// TIA Portal V19 export
DATA_BLOCK "Pumps Data"   // DB4
{ S7_Optimized_Access := 'FALSE'; DB_Accessible_From_OPC_UA := 'FALSE' }
// stored: DBAccessibleFromOPCUA false
   VAR RETAIN
      R1_CP01 : Struct
         MCMD : Bool;
         CMD : Bool;
         RESET : Bool;
         WT_SP : Time := T#5s;
         STATUS : Int;
      END_STRUCT;
      R1_AG01 : Struct
         MCMD : Bool;
         CMD : Bool;
         RESET : Bool;
         WT_SP : Time;
         STATUS : Int;
      END_STRUCT;
      CHS_CP01 : Struct
         MCMD : Bool;
         CMD : Bool;
         RESET : Bool;
         WT_SP : Time := T#5s;
         STATUS : Int;
         PUMP_SEL : Bool;
      END_STRUCT;
      CHS_CP02 : Struct
         MCMD : Bool;
         CMD : Bool;
         RESET : Bool;
         WT_SP : Time := T#5s;
         STATUS : Int;
         PUMP_SEL : Bool;
      END_STRUCT;
      CHS_CP03 : Struct
         MCMD : Bool;
         CMD : Bool;
         RESET : Bool;
         WT_SP : Time := T#5s;
         STATUS : Int;
         PUMP_SEL : Bool;
      END_STRUCT;
      R2_CP01 : Struct
         MCMD : Bool;
         CMD : Bool;
         RESET : Bool;
         WT_SP : Time := T#5s;
         STATUS : Int;
      END_STRUCT;
      R2_AG01 : Struct
         MCMD : Bool;
         CMD : Bool;
         RESET : Bool;
         WT_SP : Time;
         STATUS : Int;
      END_STRUCT;
      R3_CP01 : Struct
         MCMD : Bool;
         CMD : Bool;
         RESET : Bool;
         WT_SP : Time := T#5s;
         STATUS : Int;
      END_STRUCT;
      R3_AG01 : Struct
         MCMD : Bool;
         CMD : Bool;
         RESET : Bool;
         WT_SP : Time;
         STATUS : Int;
      END_STRUCT;
      R4_CP01 : Struct
         MCMD : Bool;
         CMD : Bool;
         RESET : Bool;
         WT_SP : Time := T#5s;
         STATUS : Int;
      END_STRUCT;
      R4_AG01 : Struct
         MCMD : Bool;
         CMD : Bool;
         RESET : Bool;
         WT_SP : Time;
         STATUS : Int;
      END_STRUCT;
      R5_CP01 : Struct
         MCMD : Bool;
         CMD : Bool;
         RESET : Bool;
         WT_SP : Time := T#5s;
         STATUS : Int;
      END_STRUCT;
      R5_AG01 : Struct
         MCMD : Bool;
         CMD : Bool;
         RESET : Bool;
         WT_SP : Time;
         STATUS : Int;
      END_STRUCT;
      R6_CP01 : Struct
         MCMD : Bool;
         CMD : Bool;
         RESET : Bool;
         WT_SP : Time := T#5s;
         STATUS : Int;
      END_STRUCT;
      R6_AG01 : Struct
         MCMD : Bool;
         CMD : Bool;
         RESET : Bool;
         WT_SP : Time;
         STATUS : Int;
      END_STRUCT;
      R7_CP01 : Struct
         MCMD : Bool;
         CMD : Bool;
         RESET : Bool;
         WT_SP : Time := T#5s;
         STATUS : Int;
      END_STRUCT;
      R7_AG01 : Struct
         MCMD : Bool;
         CMD : Bool;
         RESET : Bool;
         WT_SP : Time;
         STATUS : Int;
      END_STRUCT;
      R8_CP01 : Struct
         MCMD : Bool;
         CMD : Bool;
         RESET : Bool;
         WT_SP : Time := T#5s;
         STATUS : Int;
      END_STRUCT;
      R8_AG01 : Struct
         MCMD : Bool;
         CMD : Bool;
         RESET : Bool;
         WT_SP : Time;
         STATUS : Int;
      END_STRUCT;
      R9_CP01 : Struct
         MCMD : Bool;
         CMD : Bool;
         RESET : Bool;
         WT_SP : Time := T#5s;
         STATUS : Int;
      END_STRUCT;
      R9_AG01 : Struct
         MCMD : Bool;
         CMD : Bool;
         RESET : Bool;
         WT_SP : Time;
         STATUS : Int;
      END_STRUCT;
      R10_CP01 : Struct
         MCMD : Bool;
         CMD : Bool;
         RESET : Bool;
         WT_SP : Time := T#5s;
         STATUS : Int;
      END_STRUCT;
      R10_AG01 : Struct
         MCMD : Bool;
         CMD : Bool;
         RESET : Bool;
         WT_SP : Time;
         STATUS : Int;
      END_STRUCT;
      R11_CP01 : Struct
         MCMD : Bool;
         CMD : Bool;
         RESET : Bool;
         WT_SP : Time := T#5s;
         STATUS : Int;
      END_STRUCT;
      R11_AG01 : Struct
         MCMD : Bool;
         CMD : Bool;
         RESET : Bool;
         WT_SP : Time;
         STATUS : Int;
      END_STRUCT;
      R12_CP01 : Struct
         MCMD : Bool;
         CMD : Bool;
         RESET : Bool;
         WT_SP : Time := T#5s;
         STATUS : Int;
      END_STRUCT;
      R12_AG01 : Struct
         MCMD : Bool;
         CMD : Bool;
         RESET : Bool;
         WT_SP : Time;
         STATUS : Int;
      END_STRUCT;
      R13_CP01 : Struct
         MCMD : Bool;
         CMD : Bool;
         RESET : Bool;
         WT_SP : Time := T#5s;
         STATUS : Int;
      END_STRUCT;
      R13_AG01 : Struct
         MCMD : Bool;
         CMD : Bool;
         RESET : Bool;
         WT_SP : Time;
         STATUS : Int;
      END_STRUCT;
      R14_CP01 : Struct
         MCMD : Bool;
         CMD : Bool;
         RESET : Bool;
         WT_SP : Time := T#5s;
         STATUS : Int;
      END_STRUCT;
      R14_AG01 : Struct
         MCMD : Bool;
         CMD : Bool;
         RESET : Bool;
         WT_SP : Time;
         STATUS : Int;
      END_STRUCT;
      R15_CP01 : Struct
         MCMD : Bool;
         CMD : Bool;
         RESET : Bool;
         WT_SP : Time := T#5s;
         STATUS : Int;
      END_STRUCT;
      R15_AG01 : Struct
         MCMD : Bool;
         CMD : Bool;
         RESET : Bool;
         WT_SP : Time;
         STATUS : Int;
      END_STRUCT;
      R16_CP01 : Struct
         MCMD : Bool;
         CMD : Bool;
         RESET : Bool;
         WT_SP : Time := T#5s;
         STATUS : Int;
      END_STRUCT;
      R16_AG01 : Struct
         MCMD : Bool;
         CMD : Bool;
         RESET : Bool;
         WT_SP : Time;
         STATUS : Int;
      END_STRUCT;
      R17_CP01 : Struct
         MCMD : Bool;
         CMD : Bool;
         RESET : Bool;
         WT_SP : Time := T#5s;
         STATUS : Int;
      END_STRUCT;
      R17_AG01 : Struct
         MCMD : Bool;
         CMD : Bool;
         RESET : Bool;
         WT_SP : Time;
         STATUS : Int;
      END_STRUCT;
      R18_CP01 : Struct
         MCMD : Bool;
         CMD : Bool;
         RESET : Bool;
         WT_SP : Time := T#5s;
         STATUS : Int;
      END_STRUCT;
      R18_AG01 : Struct
         MCMD : Bool;
         CMD : Bool;
         RESET : Bool;
         WT_SP : Time;
         STATUS : Int;
      END_STRUCT;
      UCHS_CP01 : Struct
         MCMD : Bool;
         CMD : Bool;
         RESET : Bool;
         WT_SP : Time := T#5s;
         STATUS : Int;
         PUMP_SEL : Bool;
      END_STRUCT;
      UCHS_CP02 : Struct
         MCMD : Bool;
         CMD : Bool;
         RESET : Bool;
         WT_SP : Time := T#5s;
         STATUS : Int;
         PUMP_SEL : Bool;
      END_STRUCT;
      UCHS_PUPM_FAULT : Struct
         UCHS_CP01_FAIL_TO_RUN : Bool;
         UCHS_CP02_FAIL_TO_RUN : Bool;
         UCHS_CP03_FAIL_TO_RUN : Bool;
         UCHS_CP01_FAULTY : Bool;
         UCHS_CP02_FAULTY : Bool;
         UCHS_CP03_FAULTY : Bool;
      END_STRUCT;
      CS_CP01 : Struct
         MCMD : Bool;
         CMD : Bool;
         RESET : Bool;
         WT_SP : Time := T#5s;
         STATUS : Int;
         PUMP_SEL : Bool;
         "FAIL TO RUN" : Bool;
      END_STRUCT;
      CS_CP02 : Struct
         MCMD : Bool;
         CMD : Bool;
         RESET : Bool;
         WT_SP : Time := T#5s;
         STATUS : Int;
         PUMP_SEL : Bool;
         "FAIL TO RUN" : Bool;
      END_STRUCT;
      CS_CP03 : Struct
         MCMD : Bool;
         CMD : Bool;
         RESET : Bool;
         WT_SP : Time := T#5s;
         STATUS : Int;
         PUMP_SEL : Bool;
         "FAIL TO RUN" : Bool;
      END_STRUCT;
      CS_PUPM_FAULT : Struct
         CS_CP01_FAIL_TO_RUN : Bool;
         CS_CP02_FAIL_TO_RUN : Bool;
         CS_CP03_FAIL_TO_RUN : Bool;
         CS_CP01_FAULTY : Bool;
         CS_CP02_FAULTY : Bool;
         CS_CP03_FAULTY : Bool;
      END_STRUCT;
      HS_CP01 : Struct
         MCMD : Bool;
         CMD : Bool;
         RESET : Bool;
         WT_SP : Time := T#5s;
         STATUS : Int;
         PUMP_SEL : Bool;
      END_STRUCT;
      HS_CP02 : Struct
         MCMD : Bool;
         CMD : Bool;
         RESET : Bool;
         WT_SP : Time := T#5s;
         STATUS : Int;
         PUMP_SEL : Bool;
      END_STRUCT;
      HS_CP03 : Struct
         MCMD : Bool;
         CMD : Bool;
         RESET : Bool;
         WT_SP : Time := T#5s;
         STATUS : Int;
         PUMP_SEL : Bool;
      END_STRUCT;
      HS_PUPM_FAULT : Struct
         HS_CP01_FAIL_TO_RUN : Bool;
         HS_CP02_FAIL_TO_RUN : Bool;
         HS_CP03_FAIL_TO_RUN : Bool;
         HS_CP01_FAULTY : Bool;
         HS_CP02_FAULTY : Bool;
         HS_CP03_FAULTY : Bool;
      END_STRUCT;
      "A/SCRB_001_CP01" : Struct
         MCMD : Bool;
         CMD : Bool;
         RESET : Bool;
         WT_SP : Time := T#5s;
         STATUS : Int;
         PUMP_SEL : Bool;
      END_STRUCT;
      "A/SCRB_001_CP02" : Struct
         MCMD : Bool;
         CMD : Bool;
         RESET : Bool;
         WT_SP : Time := T#5s;
         STATUS : Int;
         PUMP_SEL : Bool;
      END_STRUCT;
      "A/SCRB_002_CP01" : Struct
         MCMD : Bool;
         CMD : Bool;
         RESET : Bool;
         WT_SP : Time := T#5s;
         STATUS : Int;
         PUMP_SEL : Bool;
      END_STRUCT;
      "A/SCRB_002_CP02" : Struct
         MCMD : Bool;
         CMD : Bool;
         RESET : Bool;
         WT_SP : Time := T#5s;
         STATUS : Int;
         PUMP_SEL : Bool;
      END_STRUCT;
      "A/SCRB_FAULT" : Struct
         "A/SCRB_001_CP01_FAIL_TO_RUN" : Bool;
         "A/SCRB_001_CP02_FAIL_TO_RUN" : Bool;
         "A/SCRB_002_CP01_FAIL_TO_RUN" : Bool;
         "A/SCRB_002_CP02_FAIL_TO_RUN" : Bool;
         "A/SCRB_001_BL01_FAIL_TO_RUN" : Bool;
         "A/SCRB_002_BL02_FAIL_TO_RUN" : Bool;
         "A/SCRB_001_CP01_FAULTY" : Bool;
         "A/SCRB_001_CP02_FAULTY" : Bool;
         "A/SCRB_002_CP01_FAULTY" : Bool;
         "A/SCRB_002_CP02_FAULTY" : Bool;
         "A/SCRB_001_BL01_FAULTY" : Bool;
         "A/SCRB_002_BL02_FAULTY" : Bool;
      END_STRUCT;
      "A/SCRB_001_BL01" : Struct
         MCMD : Bool;
         CMD : Bool;
         RESET : Bool;
         WT_SP : Time := T#5s;
         STATUS : Int;
         PUMP_SEL : Bool;
      END_STRUCT;
      "A/SCRB_002_BL02" : Struct
         MCMD : Bool;
         CMD : Bool;
         RESET : Bool;
         WT_SP : Time := T#5s;
         STATUS : Int;
         PUMP_SEL : Bool;
      END_STRUCT;
      "A/VP_01_CP01" : Struct
         MCMD : Bool;
         CMD : Bool;
         RESET : Bool;
         WT_SP : Time := T#5s;
         STATUS : Int;
         PUMP_SEL : Bool;
         FAULTY : Bool;
         FTR : Bool;
      END_STRUCT;
      "A/VP_02_CP01" : Struct
         MCMD : Bool;
         CMD : Bool;
         RESET : Bool;
         WT_SP : Time := T#5s;
         STATUS : Int;
         PUMP_SEL : Bool;
         FAULTY : Bool;
         FTR : Bool;
      END_STRUCT;
   END_VAR
BEGIN
END_DATA_BLOCK
